Fanuc KAREL source: KC00005.KL

PROGRAM KC00005
%NOLOCKGROUP
%ENVIRONMENT PC
VAR
  I: INTEGER
  J: INTEGER
  K: INTEGER
  R: REAL
  B: BOOLEAN
  S: STRING[80]
  T: STRING[80]
  P: PATH
  Q: PATH
  AI: ARRAY[8] OF INTEGER
  AB: ARRAY[244] OF BYTE
BEGIN
  SEND_DATAPC(I,AB,J)
END KC00005
